(* IEC 61131-3 sources: llm-plc-st-eval/data/definitivo/claude-sonnet-4-6/B8/few_shot, 3 files *)

(* ---- ejec_1.st ---- *)
```pascal
FUNCTION_BLOCK FB_Puerta
VAR_INPUT
    puertaAbierta : BOOL; (* Señal de puerta abierta *)
    reset         : BOOL; (* Reset del registro *)
END_VAR
VAR_OUTPUT
    aviso      : BOOL; (* Aviso por 5 o mas aperturas *)
    nAperturas : INT;  (* Contador de aperturas *)
END_VAR
VAR
    rTrigPuerta : R_TRIG; (* Detector de flanco ascendente *)
END_VAR

(* Detectar flanco ascendente de puertaAbierta *)
rTrigPuerta(CLK := puertaAbierta);

(* Reset tiene prioridad sobre el conteo *)
IF reset THEN
    nAperturas := 0;
ELSIF rTrigPuerta.Q THEN
    (* Incrementar solo en cada nueva apertura *)
    nAperturas := nAperturas + 1;
END_IF;

(* Activar aviso al alcanzar 5 o mas aperturas *)
aviso := nAperturas >= 5;

END_FUNCTION_BLOCK
```

(* ---- ejec_2.st ---- *)
```pascal
FUNCTION_BLOCK FB_Puerta
VAR_INPUT
    puertaAbierta : BOOL; (* Señal de puerta abierta *)
    reset         : BOOL; (* Reset del registro *)
END_VAR
VAR_OUTPUT
    aviso      : BOOL; (* Aviso por 5 o mas aperturas *)
    nAperturas : INT;  (* Contador de aperturas *)
END_VAR
VAR
    rTrigPuerta : R_TRIG; (* Detector de flanco ascendente *)
END_VAR

(* Detectar flanco ascendente de puertaAbierta *)
rTrigPuerta(CLK := puertaAbierta);

(* Reset tiene prioridad sobre el conteo *)
IF reset THEN
    nAperturas := 0;
ELSIF rTrigPuerta.Q THEN
    (* Incrementar solo en cada nueva apertura *)
    nAperturas := nAperturas + 1;
END_IF;

(* Activar aviso al alcanzar 5 o mas aperturas *)
aviso := nAperturas >= 5;

END_FUNCTION_BLOCK
```

(* ---- ejec_3.st ---- *)
```pascal
FUNCTION_BLOCK FB_Puerta
VAR_INPUT
    puertaAbierta : BOOL; (* Señal de puerta abierta *)
    reset         : BOOL; (* Pone el registro en cero *)
END_VAR
VAR_OUTPUT
    aviso      : BOOL; (* Aviso al acumular 5 o mas aperturas *)
    nAperturas : INT;  (* Contador de aperturas *)
END_VAR
VAR
    rTrigPuerta : R_TRIG; (* Detector de flanco ascendente de la puerta *)
END_VAR

(* Detectar flanco ascendente: solo cuenta la transicion FALSE->TRUE *)
rTrigPuerta(CLK := puertaAbierta);

IF reset THEN
    (* Reset: pone el contador en cero y desactiva el aviso *)
    nAperturas := 0;
ELSIF rTrigPuerta.Q THEN
    (* Nueva apertura detectada: incrementar contador *)
    nAperturas := nAperturas + 1;
END_IF;

(* Activar aviso si se han acumulado 5 o mas aperturas *)
aviso := nAperturas >= 5;
END_FUNCTION_BLOCK
```
